FUNCTION F_FeedIdString : STRING(20)
VAR_INPUT
    nFeedId : INT;
END_VAR

IF (nFeedId >= 1) AND (nFeedId <= GVL_Param.FEED_COUNT) THEN
    F_FeedIdString := GVL_Config.aFeeds[nFeedId].sId;
ELSE
    F_FeedIdString := '';
END_IF

END_FUNCTION

(* stored: Version 1.1.0.1
   POU F_FeedIdString: Id {fcb21c3a-e317-4aac-934e-ad5a53bde315}, SpecialFunc None *)
